// TIA Portal V21 export
// export: Created 2026-08-21T20:18:53.4681531Z, ExportSetting None, DisplayName Totally Integrated Automation Portal, DisplayVersion V21, DisplayName STEP 7 Professional, DisplayVersion V21, DisplayName STEP 7 Safety, DisplayVersion V21, DisplayName Tech WebApplication, DisplayVersion V21, DisplayName WinCC Basic/Comfort/Advanced, DisplayVersion V21, DisplayName WinCC Professional, DisplayVersion V21, DisplayName WinCC Unified, DisplayVersion V21
FUNCTION "Level_Sim" : Void   // FC1, FBD
{ S7_Optimized_Access := 'TRUE' }
// stored: SetENOAutomatically false
   VAR_TEMP   // added for the SCL form of the ladder/FBD networks
      _w1 : Bool;
   END_VAR
BEGIN

REGION Network 1: LevelSimulation
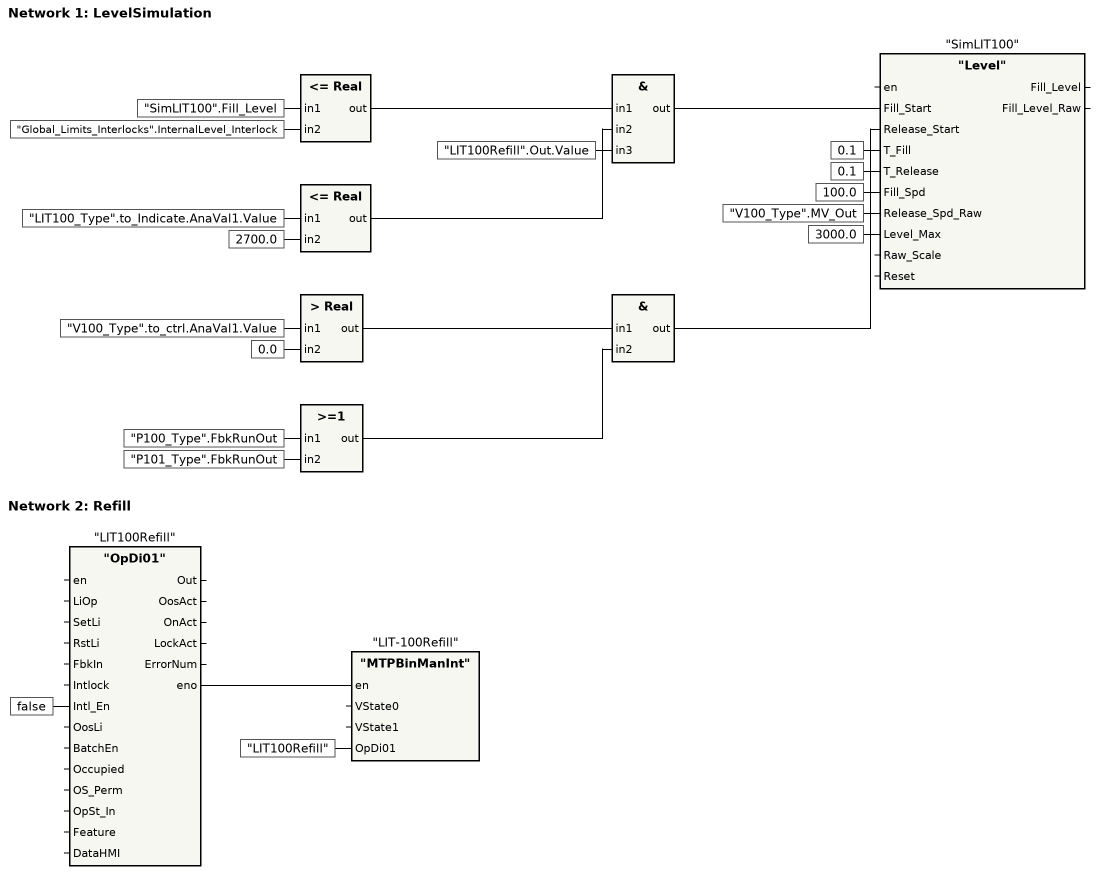
   "SimLIT100"(Fill_Start := ("SimLIT100".Fill_Level <= "Global_Limits_Interlocks".InternalLevel_Interlock) AND ("LIT100_Type".to_Indicate.AnaVal1.Value <= 2700.0) AND "LIT100Refill".Out.Value,   // "Level"
               Release_Start := ("V100_Type".to_ctrl.AnaVal1.Value > 0.0) AND ("P100_Type".FbkRunOut OR "P101_Type".FbkRunOut),
               T_Fill := 0.1,
               T_Release := 0.1,
               Fill_Spd := 100.0,
               Release_Spd_Raw := "V100_Type".MV_Out,
               Level_Max := 3000.0);
END_REGION

REGION Network 2: Refill
   "LIT100Refill"(Intl_En := false, ENO => #_w1);   // "OpDi01"
   IF #_w1 THEN
       "LIT-100Refill"(OpDi01 := "LIT100Refill");   // "MTPBinManInt"
   END_IF;
END_REGION
END_FUNCTION
